// TIA Portal V20 export
FUNCTION "GIT_Testbaustein in KOP" : Void   // FC5, LAD
{ S7_Optimized_Access := 'TRUE' }
// stored: SetENOAutomatically false
BEGIN

REGION Network 1
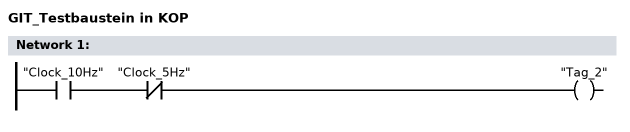
   RUNG wire#powerrail
      Contact( "Clock_10Hz" )
      I_Contact( "Clock_5Hz" )
      Coil( "Tag_2" )
   END_RUNG
   // the same network as SCL:
   "Tag_2" := "Clock_10Hz" AND NOT "Clock_5Hz";
END_REGION
END_FUNCTION
